KUKA KRL program: SplitTest2.src

&ACCESS RVP
&REL 1
&PARAM TEMPLATE = C:\KRC\Roboter\Template\vorgabe
&PARAM EDITMASK = *
DEF SplitTest2 ( )
LIN {X 549.094,Y 5.962,Z 504.960,A -174.431,B 15.001,C 175.695}
LIN {X 506.272,Y -26.320,Z 503.226,A -178.509,B 14.048,C 175.384}
LIN {X 549.094,Y 5.962,Z 504.960,A -174.431,B 15.001,C 175.695}
LIN {X 506.272,Y -26.320,Z 503.226,A -178.509,B 14.048,C 175.384}
LIN {X 549.094,Y 5.962,Z 504.960,A -174.431,B 15.001,C 175.695}
LIN {X 506.272,Y -26.320,Z 503.226,A -178.509,B 14.048,C 175.384}
LIN {X 549.094,Y 5.962,Z 504.960,A -174.431,B 15.001,C 175.695}
LIN {X 506.272,Y -26.320,Z 503.226,A -178.509,B 14.048,C 175.384}
LIN {X 549.094,Y 5.962,Z 504.960,A -174.431,B 15.001,C 175.695}
LIN {X 506.272,Y -26.320,Z 503.226,A -178.509,B 14.048,C 175.384}
LIN {X 549.094,Y 5.962,Z 504.960,A -174.431,B 15.001,C 175.695}
LIN {X 506.272,Y -26.320,Z 503.226,A -178.509,B 14.048,C 175.384}
LIN {X 549.094,Y 5.962,Z 504.960,A -174.431,B 15.001,C 175.695}
LIN {X 506.272,Y -26.320,Z 503.226,A -178.509,B 14.048,C 175.384}
LIN {X 549.094,Y 5.962,Z 504.960,A -174.431,B 15.001,C 175.695}
END
